//----------------------------------------------------------------------
// OUTPUTS TO WATCH
//----------------------------------------------------------------------
bPowered    := fbPower.Status;
bExtEnabled := fbExtEnable.Enabled;
bError      := fbPower.Error OR fbExtEnable.Error OR fbExtDisable.Error;

IF fbExtEnable.Error THEN
    nErrorID := fbExtEnable.ErrorID;
ELSIF fbPower.Error THEN
    nErrorID := fbPower.ErrorID;
ELSIF fbExtDisable.Error THEN
    nErrorID := fbExtDisable.ErrorID;
ELSE
    nErrorID := 0;
END_IF

fActPos := Axis.NcToPlc.ActPos;

END_FUNCTION_BLOCK

// ---- GlobalTextList.TcGTLO
TEXTLIST GlobalTextList
  305 = '48V  Connector Interlock'
  102 = 'Activate'
  828 = 'Battery BMS'
  548 = 'Battery BMS CMD'
  948 = 'Battery CMD'
  748 = 'Battery Control'
  71 = 'Battery Control:'
  625 = 'Battery Off'
  169 = 'Battery On'
  211 = 'Battery Relay'
  341 = 'C1 FBK'
  603 = 'C2 FBK'
  210 = 'Door monitor'
  491 = 'Door monitor solenoid'
  481 = 'Door Solenoid Status'
  551 = 'Door Status'
  131 = 'Dynamometer Safety'
  38 = 'Dynamometer Safety '
  460 = 'E.Stop - NC1'
  19 = 'E.Stop - NC2'
  512 = 'E.Stop Mentee'
  536 = 'Error'
  617 = 'Error ACK'
  361 = 'EStop Manti'
  396 = 'EStop Ok'
  665 = 'EStop1'
  338 = 'EStop2'
  865 = 'Fault / Emergency'
  954 = 'HV Connector Interlock'
  823 = 'HV Healthy'
  215 = 'HV Interlock'
  217 = 'LV Connector Interlock'
  585 = 'LV Healthy'
  227 = 'LV Interlock'
  498 = 'Mentee BOT Dynamometer'
  903 = 'Mentee BOT Dynamometer\n\tSafety '
  116 = 'Mentee BOT Dynamometer Safety '
  5 = 'Motor Cooling'
  568 = 'Motor Cooling:'
  824 = 'Open Door / Safe to Open'
  261 = 'PLC EStop'
  639 = 'RUN'
  134 = 'Run'
  727 = 'Safe to Open Door\n/ Door Opened'
  980 = 'Safety armed'
  414 = 'Safety Circut Armed'
  527 = 'Safety Circut Status'
  350 = 'Safety Refrash EStop Ok'
  97 = 'Safety Refresh\n(EStop Ok)'
  220 = 'Safety Status'
  44 = 'Safty RUN'
  830 = 'Step 1'
  699 = 'Step 2'
  745 = 'Step 3'
  789 = 'Step 4'
  483 = 'Step 5'
  652 = 'Step 6'
  264 = 'STO 1'
  577 = 'STO 2'
  298 = 'System Status'
END_TEXTLIST

// ---- VISUs/Visualization.TcVIS
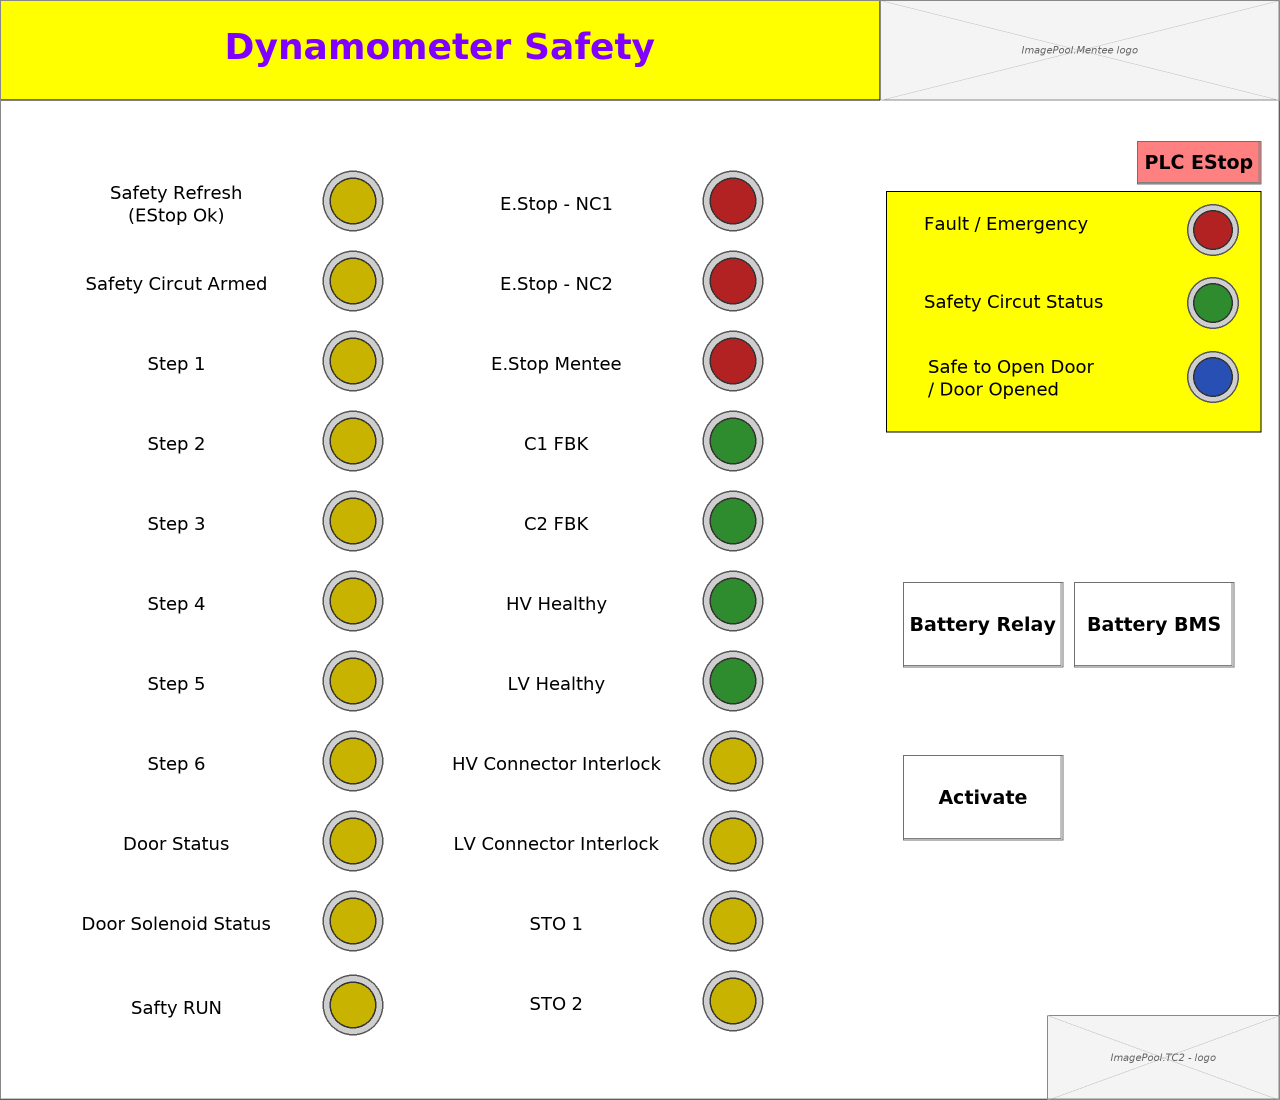
VISUALIZATION Visualization  // 1280x1100
    Rectangle (0,0 1280x1100)
    Rectangle (886,191 375x241)
    Rectangle (0,0 880x100)
    Lamp1 (318,166 70x70), variable: GVL_Safety.stTwinSAFE_IN.EStop_Ok, style: Lamp-Lamp1-Yellow
    Label (33,173 287x62), "Safety Refresh (EStop Ok)"
    Lamp1 (318,246 70x70), variable: GVL_Safety.stTwinSAFE_IN.Safety_Armed, style: Lamp-Lamp1-Yellow
    Label (33,253 287x62), "Safety Circut Armed"
    Lamp1 (318,326 70x70), variable: GVL_Safety.stTwinSAFE_IN.Speps.step1, style: Lamp-Lamp1-Yellow
    Label (33,333 287x62), "Step 1"
    Lamp1 (318,406 70x70), variable: GVL_Safety.stTwinSAFE_IN.Speps.step2, style: Lamp-Lamp1-Yellow
    Label (33,413 287x62), "Step 2"
    Lamp1 (318,486 70x70), variable: GVL_Safety.stTwinSAFE_IN.Speps.step3, style: Lamp-Lamp1-Yellow
    Label (33,493 287x62), "Step 3"
    Lamp1 (318,566 70x70), variable: GVL_Safety.stTwinSAFE_IN.Speps.step4, style: Lamp-Lamp1-Yellow
    Label (33,573 287x62), "Step 4"
    Lamp1 (318,646 70x70), variable: GVL_Safety.stTwinSAFE_IN.Speps.step5, style: Lamp-Lamp1-Yellow
    Label (33,653 287x62), "Step 5"
    Lamp1 (318,726 70x70), variable: GVL_Safety.stTwinSAFE_IN.Speps.step6, style: Lamp-Lamp1-Yellow
    Label (33,733 287x62), "Step 6"
    Lamp1 (318,806 70x70), variable: GVL_Safety.DoorMonitorFromPLC, style: Lamp-Lamp1-Yellow
    Label (33,813 287x62), "Door Status"
    Lamp1 (318,970 70x70), variable: GVL_Safety.stTwinSAFE_OUT.RUN, style: Lamp-Lamp1-Yellow
    Label (33,977 287x62), "Safty RUN"
    Lamp1 (318,886 70x70), variable: GVL_Safety.SolonoidStatus, style: Lamp-Lamp1-Yellow
    Label (33,893 287x62), "Door Solenoid Status"
    Button (1137,141 124x43), "PLC EStop", colour toggle: GVL_Safety.stTwinSAFE_OUT.EstopPLC
        toggle GVL_Safety.stTwinSAFE_OUT.EstopPLC
    Button (903,582 160x85), "Battery Relay", colour toggle: GVL_Safety.stTwinSAFE_OUT.BatRelay_CMD
        toggle GVL_Safety.stTwinSAFE_OUT.BatRelay_CMD
    Button (1074,582 160x85), "Battery BMS", colour toggle: GVL_Safety.stTwinSAFE_OUT.BatBMS_Cmd
        toggle GVL_Safety.stTwinSAFE_OUT.BatBMS_Cmd
    Lamp1 (698,166 70x70), variable: GVL_Safety.stTwinSAFE_IN.EStop_NC1, style: Lamp-Lamp1-Red
    Label (413,173 287x62), "E.Stop - NC1"
    Lamp1 (698,246 70x70), variable: GVL_Safety.stTwinSAFE_IN.EStop_NC2, style: Lamp-Lamp1-Red
    Label (413,253 287x62), "E.Stop - NC2"
    Lamp1 (698,326 70x70), variable: GVL_Safety.stTwinSAFE_IN.EStop_MantiRob, style: Lamp-Lamp1-Red
    Label (413,333 287x62), "E.Stop Mentee"
    Lamp1 (698,406 70x70), variable: GVL_Safety.stTwinSAFE_IN.C1_FBK, style: Lamp-Lamp1-Green
    Label (413,413 287x62), "C1 FBK"
    Lamp1 (698,486 70x70), variable: GVL_Safety.stTwinSAFE_IN.C2_FBK, style: Lamp-Lamp1-Green
    Label (413,493 287x62), "C2 FBK"
    Lamp1 (698,566 70x70), variable: GVL_Safety.stTwinSAFE_IN.HV_Healthy_Invert, style: Lamp-Lamp1-Green
    Label (413,573 287x62), "HV Healthy"
    Lamp1 (698,646 70x70), variable: GVL_Safety.stTwinSAFE_IN.LV_Healthy_Invert, style: Lamp-Lamp1-Green
    Label (413,653 287x62), "LV Healthy"
    Lamp1 (698,726 70x70), variable: GVL_Safety.stTwinSAFE_IN.HV_Interlock, style: Lamp-Lamp1-Yellow
    Label (413,733 287x62), "HV Connector Interlock"
    Lamp1 (698,806 70x70), variable: GVL_Safety.stTwinSAFE_IN.LV_Interlock, style: Lamp-Lamp1-Yellow
    Label (413,813 287x62), "LV Connector Interlock"
    Lamp1 (698,886 70x70), variable: GVL_Safety.stTwinSAFE_IN.STO_1, style: Lamp-Lamp1-Yellow
    Label (413,893 287x62), "STO 1"
    Lamp1 (698,966 70x70), variable: GVL_Safety.stTwinSAFE_IN.STO_2, style: Lamp-Lamp1-Yellow
    Label (413,973 287x62), "STO 2"
    Button (903,755 160x85), "Activate", colour toggle: GVL_IO.b_MotorCooling
        toggle GVL_IO.b_MotorCooling
    Image (880,0 400x100), image: ImagePool.Mentee logo
    Label (0,0 880x93), "Dynamometer Safety"
    Lamp1 (1183,200 60x60), variable: GVL_IO.RedLED, style: Lamp-Lamp1-Red
    Lamp1 (1183,273 60x60), variable: GVL_IO.GreenLED, style: Lamp-Lamp1-Green
    Lamp1 (1183,347 60x60), variable: GVL_IO.BlueLED, style: Lamp-Lamp1-Blue
    Label (921,193 195x62), "Fault / Emergency"
    Label (921,271 252x62), "Safety Circut Status"
    Label (925,347 252x62), "Safe to Open Door / Door Opened"
    Label (895,517 252x62), "Battery Control"
    Label (903,691 252x62), "Motor Cooling"
    Label (886,133 300x62), "System Status"
    Image (1047,1015 233x85), image: ImagePool.TC2 - logo
END_VISUALIZATION
